(* IEC 61131-3 sources: llm-plc-st-eval/data/calibracion/gpt-4o-2024-08-06/B1/zero_shot, 3 files *)

(* ---- ejec_1.st ---- *)
```pascal
FUNCTION_BLOCK FB_Motor
VAR_INPUT
    btnMarcha : BOOL;   // Botón de marcha
    btnParo : BOOL;     // Botón de paro
    btnEmerg : BOOL;    // Botón de paro de emergencia
END_VAR

VAR_OUTPUT
    motorOn : BOOL;     // Estado del motor (encendido/apagado)
END_VAR

VAR
    motorLatch : BOOL;  // Latch para mantener el estado del motor
    emergStopLatch : BOOL; // Latch para el estado de paro de emergencia
END_VAR

// Implementación del control de arranque y paro del motor
IF btnEmerg THEN
    // Si se presiona el botón de emergencia, activar el latch de emergencia
    emergStopLatch := TRUE;
    motorLatch := FALSE; // Apagar el motor inmediatamente
ELSIF btnParo THEN
    // Si se presiona el botón de paro, apagar el motor
    motorLatch := FALSE;
ELSIF btnMarcha AND NOT emergStopLatch THEN
    // Si se presiona el botón de marcha y no hay paro de emergencia, encender el motor
    motorLatch := TRUE;
END_IF

// Actualizar la salida del motor
motorOn := motorLatch;
```

Este código implementa el control de arranque y paro de un motor trifásico utilizando un bloque de función en Structured Text (ST). El motor se mantiene encendido al soltar el botón de marcha y se apaga al presionar el botón de paro o el de emergencia. El paro de emergencia impide que el motor vuelva a arrancar hasta que se restablezca el sistema.

(* ---- ejec_2.st ---- *)
```pascal
FUNCTION_BLOCK FB_Motor
VAR_INPUT
    btnMarcha : BOOL;   // Botón de marcha
    btnParo : BOOL;     // Botón de paro
    btnEmerg : BOOL;    // Botón de paro de emergencia
END_VAR

VAR_OUTPUT
    motorOn : BOOL;     // Estado del motor (encendido/apagado)
END_VAR

VAR
    motorLatch : BOOL;  // Latch para mantener el motor encendido
    emergStop : BOOL;   // Estado del paro de emergencia
END_VAR

// Lógica de control del motor
IF btnEmerg THEN
    // Si el botón de emergencia está presionado, apaga el motor y activa el estado de emergencia
    motorOn := FALSE;
    emergStop := TRUE;
ELSIF btnParo THEN
    // Si el botón de paro está presionado, apaga el motor
    motorOn := FALSE;
ELSE
    // Si no hay emergencia y el botón de marcha está presionado, y no hay estado de emergencia
    IF btnMarcha AND NOT emergStop THEN
        motorLatch := TRUE;  // Activa el latch del motor
    END_IF;

    // Mantiene el motor encendido si el latch está activo
    motorOn := motorLatch;
END_IF;

// Resetea el latch del motor si el motor está apagado
IF NOT motorOn THEN
    motorLatch := FALSE;
END_IF;
```

Este código implementa la lógica de control para el arranque y paro de un motor trifásico utilizando un bloque de función en Structured Text (ST). El motor se mantiene encendido mediante un latch (`motorLatch`) y se apaga al presionar el botón de paro o el de emergencia. El estado de emergencia impide el rearranque del motor hasta que se resetea.

(* ---- ejec_3.st ---- *)
```pascal
FUNCTION_BLOCK FB_Motor
VAR_INPUT
    btnMarcha : BOOL;   // Botón de marcha
    btnParo : BOOL;     // Botón de paro
    btnEmerg : BOOL;    // Botón de paro de emergencia
END_VAR

VAR_OUTPUT
    motorOn : BOOL;     // Estado del motor (encendido/apagado)
END_VAR

VAR
    motorLatch : BOOL;  // Latch para mantener el estado del motor
    emergStopLatch : BOOL; // Latch para el estado de paro de emergencia
END_VAR

// Lógica de control del motor
IF btnEmerg THEN
    // Si se presiona el botón de emergencia, activar el latch de emergencia
    emergStopLatch := TRUE;
    motorLatch := FALSE; // Apagar el motor inmediatamente
ELSIF btnParo THEN
    // Si se presiona el botón de paro, apagar el motor
    motorLatch := FALSE;
ELSIF btnMarcha AND NOT emergStopLatch THEN
    // Si se presiona el botón de marcha y no hay paro de emergencia, encender el motor
    motorLatch := TRUE;
END_IF

// Actualizar el estado de salida del motor
motorOn := motorLatch;

// Resetear el latch de emergencia si el motor está apagado
IF NOT motorLatch THEN
    emergStopLatch := FALSE;
END_IF

END_FUNCTION_BLOCK
```

Este código implementa un control básico de arranque y paro de un motor trifásico utilizando un bloque de función en Structured Text (ST) conforme al estándar IEC 61131-3. El motor se mantiene encendido después de soltar el botón de marcha y se apaga al presionar el botón de paro o el de emergencia. Además, el motor no se rearranca automáticamente después de un paro de emergencia hasta que se libere y vuelva a presionar el botón de marcha.
